TYPE stShutterState :
STRUCT
    CurrentStateType    : eShutterStateType;
    PreviousStateType   : eShutterStateType;
END_STRUCT
END_TYPE

(* stored: Version 1.1.0.1
   DUT stShutterState: Id {777aa08a-edfb-4ead-b67a-bc47756d0cde} *)
